Fanuc KAREL source: ko00062.KL

-- PROVISIONAL review KL for V1013-1; original PC SHA256 d2bddd6a16f93178917139cd9c4abd4d3a85532cf00f2923c003f8c83b27cc0a
-- Incomplete behavior may be omitted. Consult companion uncertainty JSON. Do not deploy.
PROGRAM KO00062
%NOLOCKGROUP
BEGIN
  -- UNRESOLVED_PC offsets 5-12; opcodes 9D,23
  -- UNRESOLVED_PC offsets 17-69; opcodes 27,27,49,7E,AD,27,49,7E,AD,22,31,7E,4A
  -- UNRESOLVED_PC offsets 74-78; opcodes 7F
END KO00062
